(* IEC 61131-3 sources: plc-process-lib/tests/POUs/Suites/FB_AnalogInput_Test, 80 files *)

(* ---- AlarmEventsFailureValueIsRawInput.method.decl.st ---- *)
// Номера и значения событий: udiAlarmIdBase 120 — тревога HH = 120, Failure = 124; значение события HH — rValue_eu
// (95), Failure — сырое rIn (22,5 мА).
METHOD PRIVATE AlarmEventsFailureValueIsRawInput
VAR
    fbTime : FB_FakeTime;         // подменное время
    fbAi   : FB_AnalogInput;      // ФБ под тестом
    stCmd  : ST_AnalogInputCmd;   // команды
    stCfg  : ST_AnalogInputCfg;   // конфигурация
    fbSink : FB_TestSink;         // приёмник событий
    stEv   : ST_AlarmEvent;       // событие
END_VAR

(* ---- At20p5mAIsGood.method.decl.st ---- *)
// Граница 20,5 мА — ещё норма (NE43_MEAS_HIGH_MA: «I > — вне диапазона»): Good, значение 103,125 %.
METHOD PRIVATE At20p5mAIsGood
VAR
    fbTime : FB_FakeTime;         // подменное время
    fbAi   : FB_AnalogInput;      // ФБ под тестом
    stCmd  : ST_AnalogInputCmd;   // команды
    stCfg  : ST_AnalogInputCfg;   // конфигурация
END_VAR

(* ---- At20p7mAIsOutOfSpecification.method.decl.st ---- *)
// 20,7 мА (между 20,5 и 21,0): OverRange, OutOfSpecification, значение — насыщение NE 43 20,5 мА (103,125 %), без
// экстраполяции; выход за диапазон подтверждён — xValid = FALSE (AI-13), бит AI_WRN_OVER_RANGE.
// источник: tools/reference/ai_reference.py, сценарий scale «20,7 мА, шкала 0..100 (насыщение NE 43)».
METHOD PRIVATE At20p7mAIsOutOfSpecification
VAR
    fbTime : FB_FakeTime;         // подменное время
    fbAi   : FB_AnalogInput;      // ФБ под тестом
    stCmd  : ST_AnalogInputCmd;   // команды
    stCfg  : ST_AnalogInputCfg;   // конфигурация
END_VAR

(* ---- At21mAIsFailure.method.decl.st ---- *)
// Граница NE 43 21,0 мА включена в отказ (A-02): FailHigh, Failure, бит AI_FLT_FAIL_HIGH; 20,99 мА — ещё OverRange.
METHOD PRIVATE At21mAIsFailure
VAR
    fbTime : FB_FakeTime;         // подменное время
    fbAi   : FB_AnalogInput;      // ФБ под тестом
    stCmd  : ST_AnalogInputCmd;   // команды
    stCfg  : ST_AnalogInputCfg;   // конфигурация
END_VAR

(* ---- At3p6mAIsFailure.method.decl.st ---- *)
// Граница NE 43 3,6 мА включена в отказ (A-02, сверить с NAMUR NE 43): FailLow, Failure (tFailDelay = 0), бит
// AI_FLT_FAIL_LOW; чуть выше, 3,61 мА — уже UnderRange.
METHOD PRIVATE At3p6mAIsFailure
VAR
    fbTime : FB_FakeTime;         // подменное время
    fbAi   : FB_AnalogInput;      // ФБ под тестом
    stCmd  : ST_AnalogInputCmd;   // команды
    stCfg  : ST_AnalogInputCfg;   // конфигурация
END_VAR

(* ---- At3p7mAIsOutOfSpecification.method.decl.st ---- *)
// 3,7 мА (между 3,6 и 3,8): UnderRange, OutOfSpecification, значение — насыщение NE 43 3,8 мА (-1,25 %), без
// экстраполяции; выход за диапазон подтверждён (tFailDelay = 0) — xValid = FALSE (AI-13), бит AI_WRN_UNDER_RANGE,
// тревога OutOfRange. источник: tools/reference/ai_reference.py, сценарий scale «3,7 мА, шкала 0..100 (насыщение
// NE 43)».
METHOD PRIVATE At3p7mAIsOutOfSpecification
VAR
    fbTime : FB_FakeTime;         // подменное время
    fbAi   : FB_AnalogInput;      // ФБ под тестом
    stCmd  : ST_AnalogInputCmd;   // команды
    stCfg  : ST_AnalogInputCfg;   // конфигурация
    itfAlm : I_Alarm;             // слот тревоги через интерфейс
END_VAR

(* ---- At3p8mAIsGood.method.decl.st ---- *)
// Граница 3,8 мА — уже норма (NE43_MEAS_LOW_MA: «I < — вне диапазона»): Good, значение -1,25 %.
METHOD PRIVATE At3p8mAIsGood
VAR
    fbTime : FB_FakeTime;         // подменное время
    fbAi   : FB_AnalogInput;      // ФБ под тестом
    stCmd  : ST_AnalogInputCmd;   // команды
    stCfg  : ST_AnalogInputCfg;   // конфигурация
END_VAR

(* ---- CfgErrBitsMatchContractMap.method.decl.st ---- *)
// Каждая проверка CheckConfig ставит свой бит wCfgErr (карта 11.5): тип входа вне перечисления, шкала, порядок уставок,
// уставка вне шкалы, гистерезис (< 0 и >= диапазона), отсечка (вне 0…20 %), значение отказа (вне перечисления и NaN),
// приоритет тревоги вне перечисления, шкала отсчётов Raw. Один экземпляр: wCfgErr — результат проверки этого вызова.
METHOD PRIVATE CfgErrBitsMatchContractMap
VAR
    fbTime : FB_FakeTime;         // подменное время
    fbAi   : FB_AnalogInput;      // ФБ под тестом
    stCmd  : ST_AnalogInputCmd;   // команды
    stCfg  : ST_AnalogInputCfg;   // конфигурация
    stBad  : ST_AnalogInputCfg;   // испорченная копия
    uEnum  : U_AiDiTestEnum;      // значение вне строгого перечисления
    uPrio  : U_TestEnumInt;       // приоритет вне перечисления
    uBits  : U_RealBits;          // NaN по битам
END_VAR

(* ---- ChannelFaultSetsFailure.method.decl.st ---- *)
// xChannelFault (диагностика модуля, ошибка обмена) при нормальном токе: ChannelFault, значение удерживается, через
// tFailDelay 2 с — Failure и бит AI_FLT_CHANNEL; после снятия — возврат через те же 2 с.
METHOD PRIVATE ChannelFaultSetsFailure
VAR
    fbTime : FB_FakeTime;         // подменное время
    fbAi   : FB_AnalogInput;      // ФБ под тестом
    stCmd  : ST_AnalogInputCmd;   // команды
    stCfg  : ST_AnalogInputCfg;   // конфигурация
    iStep  : INT;                 // шаг цикла
END_VAR

(* ---- ChannelFaultSetsFailure.method.impl.st ---- *)
coUnit.TEST('AnalogInput_ChannelFault_SetsFailure');

fbAi(itfTime := fbTime, rIn := 12.0, stCmd := stCmd, stCfg := stCfg);   // t0: 50
fbTime.Advance(tStep := T#100MS);
// t1 = t0 + 0,1 с: отказ канала
fbAi(itfTime := fbTime, rIn := 12.0, xChannelFault := TRUE, stCmd := stCmd, stCfg := stCfg);
FOR iStep := 1 TO 19 DO   // t1 + 1,9 с
    fbTime.Advance(tStep := T#100MS);
    fbAi(itfTime := fbTime, rIn := 12.0, xChannelFault := TRUE, stCmd := stCmd, stCfg := stCfg);
END_FOR
AssertTrue(Condition := fbAi.stSts.eSignal = E_AiSignalState.ChannelFault, Message := 'ChannelFault');
AssertFalse(Condition := fbAi.Fault, Message := 'no failure before tFailDelay');
fbTime.Advance(tStep := T#100MS);
fbAi(itfTime := fbTime, rIn := 12.0, xChannelFault := TRUE, stCmd := stCmd, stCfg := stCfg);   // t1 + 2,0 с
AssertTrue(Condition := fbAi.Fault, Message := 'failure after tFailDelay');
AssertEquals_WORD(Expected := GVL_Const.AI_FLT_CHANNEL, Actual := fbAi.stSts.stCommon.wFault, Message := 'CHANNEL bit');
AssertEquals_REAL(Expected := 50.0, Actual := fbAi.rValue_eu, Delta := 1.0E-4, Message := 'value held');
fbTime.Advance(tStep := T#100MS);
fbAi(itfTime := fbTime, rIn := 12.0, xChannelFault := FALSE, stCmd := stCmd, stCfg := stCfg);   // tc: отказ канала снят
FOR iStep := 1 TO 19 DO   // tc + 1,9 с
    fbTime.Advance(tStep := T#100MS);
    fbAi(itfTime := fbTime, rIn := 12.0, xChannelFault := FALSE, stCmd := stCmd, stCfg := stCfg);
END_FOR
AssertTrue(Condition := fbAi.Fault, Message := 'failure kept during return confirmation');
AssertEquals_WORD(Expected := 0, Actual := fbAi.stSts.stCommon.wFault,
                  Message := 'fault bit by current classification');
FOR iStep := 1 TO 1 DO   // tc + 2,0 с
    fbTime.Advance(tStep := T#100MS);
    fbAi(itfTime := fbTime, rIn := 12.0, xChannelFault := FALSE, stCmd := stCmd, stCfg := stCfg);
END_FOR
AssertFalse(Condition := fbAi.Fault, Message := 'failure cleared');

coUnit.TEST_FINISHED();

(* ---- ClampLimitsToRange.method.decl.st ---- *)
// По умолчанию значение экстраполируется (20,4 мА — 102,5 %); с xClamp — ограничено шкалой (100 и 0) с предупреждением
// AI_WRN_CLAMPED. источник: tools/reference/ai_reference.py, сценарии scale «20,4 мА без ограничения», «… с
// ограничением», «3,9 мА с ограничением».
METHOD PRIVATE ClampLimitsToRange
VAR
    fbTime : FB_FakeTime;         // подменное время
    fbAi   : FB_AnalogInput;      // ФБ под тестом
    stCmd  : ST_AnalogInputCmd;   // команды
    stCfg  : ST_AnalogInputCfg;   // конфигурация
END_VAR

(* ---- DefaultCfgFirstCallAutoTypeAndSlots.method.decl.st ---- *)
// Cfg по умолчанию проходит CheckConfig (wCfgErr = 0); после первого вызова — Auto («Измерение»), тип AnalogInput, 6
// слотов тревог, Good, бит DEV_STS_MODE_AUTO; седьмого слота нет; Local не запрашивается.
METHOD PRIVATE DefaultCfgFirstCallAutoTypeAndSlots
VAR
    fbTime : FB_FakeTime;         // подменное время
    fbAi   : FB_AnalogInput;      // ФБ под тестом
    stCmd  : ST_AnalogInputCmd;   // команды
    stCfg  : ST_AnalogInputCfg;   // конфигурация
    itfAlm : I_Alarm;             // слот тревоги через интерфейс
END_VAR

(* ---- EngInputPassesThrough.method.decl.st ---- *)
// Eng (значение уже в инж. ед., Modbus REAL): шкала -50..150, 123,4 — 123,4 (86,7 %); NE 43 не применяется (0 — норма).
// источник: tools/reference/ai_reference.py, сценарий scale «Eng 123,4, шкала -50..150».
METHOD PRIVATE EngInputPassesThrough
VAR
    fbTime : FB_FakeTime;         // подменное время
    fbAi   : FB_AnalogInput;      // ФБ под тестом
    stCmd  : ST_AnalogInputCmd;   // команды
    stCfg  : ST_AnalogInputCfg;   // конфигурация
END_VAR

(* ---- FailureForcesLimitsFalseAndSuppressesLimitAlarms.method.decl.st ---- *)
// H 4,0 активна (4,25 м); обрыв: пока отказ не подтверждён, H держится по удержанному значению, ложного LL (0,5) нет;
// после подтверждения флаги сняты, тревога H — SuppressedByDesign, тревога Failure — ActiveUnack.
METHOD PRIVATE FailureForcesLimitsFalseAndSuppressesLimitAlarms
VAR
    fbTime : FB_FakeTime;         // подменное время
    fbAi   : FB_AnalogInput;      // ФБ под тестом
    stCmd  : ST_AnalogInputCmd;   // команды
    stCfg  : ST_AnalogInputCfg;   // конфигурация
    itfAlm : I_Alarm;             // слот тревоги через интерфейс
    iStep  : INT;                 // шаг цикла
END_VAR

(* ---- FailureForcesLimitsFalseAndSuppressesLimitAlarms.method.impl.st ---- *)
coUnit.TEST('AnalogInput_Failure_ForcesLimitsFalseAndSuppressesLimitAlarms');

stCfg.rRangeHi_eu := 5.0;
SetLimit(stCfgAi := stCfg, uiIdx := E_AiAlarm.H, xEnable := TRUE, rSp_eu := 4.0, rHyst_eu := 0.1, tOnDly := T#0S,
         tOffDly := T#0S);
SetLimit(stCfgAi := stCfg, uiIdx := E_AiAlarm.LL, xEnable := TRUE, rSp_eu := 0.5, rHyst_eu := 0.1, tOnDly := T#0S,
         tOffDly := T#0S);
fbAi(itfTime := fbTime, rIn := 17.6, stCmd := stCmd, stCfg := stCfg);   // t0: 4,25 м
AssertTrue(Condition := fbAi.xH, Message := 'H active before break');
itfAlm := fbAi.GetAlarm(uiIndex := E_AiAlarm.H);
AssertTrue(Condition := itfAlm.State = E_AlarmState.ActiveUnack, Message := 'H alarm active');
fbTime.Advance(tStep := T#100MS);
fbAi(itfTime := fbTime, rIn := 0.0, stCmd := stCmd, stCfg := stCfg);   // t1 = t0 + 0,1 с: обрыв
FOR iStep := 1 TO 19 DO   // t1 + 1,9 с
    fbTime.Advance(tStep := T#100MS);
    fbAi(itfTime := fbTime, rIn := 0.0, stCmd := stCmd, stCfg := stCfg);
END_FOR
AssertTrue(Condition := fbAi.xH, Message := 'H kept on held value while pending');
AssertFalse(Condition := fbAi.xLL, Message := 'no false LL while pending');
fbTime.Advance(tStep := T#100MS);
fbAi(itfTime := fbTime, rIn := 0.0, stCmd := stCmd, stCfg := stCfg);   // t1 + 2,0 с
AssertTrue(Condition := fbAi.Fault, Message := 'failure confirmed');
AssertFalse(Condition := fbAi.xH, Message := 'H forced off');
AssertFalse(Condition := fbAi.xLL, Message := 'LL forced off');
AssertTrue(Condition := itfAlm.State = E_AlarmState.SuppressedByDesign, Message := 'H alarm suppressed');
itfAlm := fbAi.GetAlarm(uiIndex := E_AiAlarm.Failure);
AssertTrue(Condition := itfAlm.State = E_AlarmState.ActiveUnack, Message := 'failure alarm');

coUnit.TEST_FINISHED();

(* ---- FailValueSubstituteUsesCfgValue.method.decl.st ---- *)
// eFailValue = Substitute: до подтверждения отказа держится последнее хорошее значение (25), после — rFailValue_eu =
// 99, xValid = FALSE.
METHOD PRIVATE FailValueSubstituteUsesCfgValue
VAR
    fbTime : FB_FakeTime;         // подменное время
    fbAi   : FB_AnalogInput;      // ФБ под тестом
    stCmd  : ST_AnalogInputCmd;   // команды
    stCfg  : ST_AnalogInputCfg;   // конфигурация
    iStep  : INT;                 // шаг цикла
END_VAR

(* ---- FailValueSubstituteUsesCfgValue.method.impl.st ---- *)
coUnit.TEST('AnalogInput_FailValueSubstitute_UsesCfgValue');

stCfg.eFailValue := E_AiFailValue.Substitute;
stCfg.rFailValue_eu := 99.0;
stCfg.tFailDelay := T#1S;
fbAi(itfTime := fbTime, rIn := 8.0, stCmd := stCmd, stCfg := stCfg);   // t0: 25
fbTime.Advance(tStep := T#100MS);
fbAi(itfTime := fbTime, rIn := 0.0, stCmd := stCmd, stCfg := stCfg);   // t1 = t0 + 0,1 с: обрыв
FOR iStep := 1 TO 9 DO   // t1 + 0,9 с
    fbTime.Advance(tStep := T#100MS);
    fbAi(itfTime := fbTime, rIn := 0.0, stCmd := stCmd, stCfg := stCfg);
END_FOR
AssertEquals_REAL(Expected := 25.0, Actual := fbAi.rValue_eu, Delta := 1.0E-4, Message := 'last good while pending');
AssertTrue(Condition := fbAi.xValid, Message := 'valid while pending');
FOR iStep := 1 TO 1 DO   // t1 + 1,0 с
    fbTime.Advance(tStep := T#100MS);
    fbAi(itfTime := fbTime, rIn := 0.0, stCmd := stCmd, stCfg := stCfg);
END_FOR
AssertTrue(Condition := fbAi.Fault, Message := 'failure confirmed');
AssertEquals_REAL(Expected := 99.0, Actual := fbAi.rValue_eu, Delta := 0.0, Message := 'substitute value from Cfg');
AssertFalse(Condition := fbAi.xValid, Message := 'substitute value is not valid');

coUnit.TEST_FINISHED();

(* ---- FilterIndependentOfCycleTime.method.decl.st ---- *)
// Один и тот же интервал 5 с при T = 10 с: шаг 10 мс (500 вызовов), 250 мс (20 вызовов) и неравномерный 50/150/300 мс
// дают одно значение 39,347 (1 - e^-0,5): фильтр считает по реальному шагу времени. Неявный Эйлер dt/(T + dt) при 250
// мс дал бы 38,97. источник: tools/reference/ai_reference.py, сценарии filter «5 с шагом 10 мс», «… 250 мс», «…
// неравномерно».
METHOD PRIVATE FilterIndependentOfCycleTime
VAR
    fbTimeA : FB_FakeTime;         // время экземпляра A
    fbTimeB : FB_FakeTime;         // время экземпляра B
    fbTimeC : FB_FakeTime;         // время экземпляра C
    fbAiA   : FB_AnalogInput;      // шаг 10 мс
    fbAiB   : FB_AnalogInput;      // шаг 250 мс
    fbAiC   : FB_AnalogInput;      // неравномерный шаг
    stCmdA  : ST_AnalogInputCmd;   // команды A
    stCmdB  : ST_AnalogInputCmd;   // команды B
    stCmdC  : ST_AnalogInputCmd;   // команды C
    stCfg   : ST_AnalogInputCfg;   // конфигурация
    iStep   : INT;                 // шаг цикла
END_VAR

(* ---- FilterIndependentOfCycleTime.method.impl.st ---- *)
coUnit.TEST('AnalogInput_Filter_IndependentOfCycleTime');

stCfg.tFilter := T#10S;
fbAiA(itfTime := fbTimeA, rIn := 4.0, stCmd := stCmdA, stCfg := stCfg);
fbAiB(itfTime := fbTimeB, rIn := 4.0, stCmd := stCmdB, stCfg := stCfg);
fbAiC(itfTime := fbTimeC, rIn := 4.0, stCmd := stCmdC, stCfg := stCfg);
FOR iStep := 1 TO 500 DO
    fbTimeA.Advance(tStep := T#10MS);
    fbAiA(itfTime := fbTimeA, rIn := 20.0, stCmd := stCmdA, stCfg := stCfg);
END_FOR
FOR iStep := 1 TO 20 DO
    fbTimeB.Advance(tStep := T#250MS);
    fbAiB(itfTime := fbTimeB, rIn := 20.0, stCmd := stCmdB, stCfg := stCfg);
END_FOR
FOR iStep := 1 TO 10 DO
    fbTimeC.Advance(tStep := T#50MS);
    fbAiC(itfTime := fbTimeC, rIn := 20.0, stCmd := stCmdC, stCfg := stCfg);
    fbTimeC.Advance(tStep := T#150MS);
    fbAiC(itfTime := fbTimeC, rIn := 20.0, stCmd := stCmdC, stCfg := stCfg);
    fbTimeC.Advance(tStep := T#300MS);
    fbAiC(itfTime := fbTimeC, rIn := 20.0, stCmd := stCmdC, stCfg := stCfg);
END_FOR
AssertEquals_REAL(Expected := 39.34694, Actual := fbAiA.rValue_eu, Delta := 1.0E-3, Message := '10 ms steps');
AssertEquals_REAL(Expected := 39.34694, Actual := fbAiB.rValue_eu, Delta := 1.0E-3, Message := '250 ms steps');
AssertEquals_REAL(Expected := 39.34694, Actual := fbAiC.rValue_eu, Delta := 1.0E-3, Message := 'irregular steps');
AssertEquals_REAL(Expected := fbAiA.rValue_eu, Actual := fbAiB.rValue_eu, Delta := 1.0E-4,
                  Message := 'same result for 10 ms and 250 ms');

coUnit.TEST_FINISHED();

(* ---- FilterOneTimeConstantReaches63Pct.method.decl.st ---- *)
// Фильтр T = 10 с, ступень 0 -> 100 % с шагом 100 мс: в 9,9 с — 62,842, ровно через T — 63,212 (1 - e^-1). источник:
// tools/reference/ai_reference.py, сценарии filter «… 99 шагов по 0,1 с» и «… 100 шагов по 0,1 с».
METHOD PRIVATE FilterOneTimeConstantReaches63Pct
VAR
    fbTime : FB_FakeTime;         // подменное время
    fbAi   : FB_AnalogInput;      // ФБ под тестом
    stCmd  : ST_AnalogInputCmd;   // команды
    stCfg  : ST_AnalogInputCfg;   // конфигурация
    iStep  : INT;                 // шаг цикла
END_VAR

(* ---- FilterOneTimeConstantReaches63Pct.method.impl.st ---- *)
coUnit.TEST('AnalogInput_Filter_OneTimeConstant_Reaches63Pct');

stCfg.tFilter := T#10S;
fbAi(itfTime := fbTime, rIn := 4.0, stCmd := stCmd, stCfg := stCfg);   // t0: фильтр начат с 0
FOR iStep := 1 TO 99 DO   // ступень 100 %, t0 + 9,9 с
    fbTime.Advance(tStep := T#100MS);
    fbAi(itfTime := fbTime, rIn := 20.0, stCmd := stCmd, stCfg := stCfg);
END_FOR
AssertEquals_REAL(Expected := 62.84233, Actual := fbAi.rValue_eu, Delta := 1.0E-3, Message := '62.84 at 9.9 s');
fbTime.Advance(tStep := T#100MS);
fbAi(itfTime := fbTime, rIn := 20.0, stCmd := stCmd, stCfg := stCfg);   // t0 + 10,0 с
AssertEquals_REAL(Expected := 63.21206, Actual := fbAi.rValue_eu, Delta := 1.0E-3, Message := '63.2 % after one T');

coUnit.TEST_FINISHED();

(* ---- GuardBandHighInvalidLimitsKept.method.decl.st ---- *)
// 20,9 мА — верхняя защитная полоса NE 43 (между 20,5 и 21 мА, AI-13): значение — насыщение 20,5 мА, 10,3125 м на
// шкале 0..10 м (1,03125 · 10), без экстраполяции; через tFailDelay — xValid = FALSE, OVER_RANGE, уставка HH (9,5 м)
// остаётся: процесс выше верхнего предела измерения. источник: tools/reference/ai_reference.py, сценарий scale
// «20,9 мА, шкала 0..10 (насыщение NE 43)».
METHOD PRIVATE GuardBandHighInvalidLimitsKept
VAR
    fbTime : FB_FakeTime;         // подменное время
    fbAi   : FB_AnalogInput;      // ФБ под тестом
    stCmd  : ST_AnalogInputCmd;   // команды
    stCfg  : ST_AnalogInputCfg;   // конфигурация
    iStep  : INT;                 // шаг цикла
END_VAR

(* ---- GuardBandHighInvalidLimitsKept.method.impl.st ---- *)
coUnit.TEST('AnalogInput_GuardBandHigh_InvalidLimitsKept');

stCfg.rRangeHi_eu := 10.0;
stCfg.astLimit[E_AiAlarm.HH].xEnable := TRUE;
stCfg.astLimit[E_AiAlarm.HH].rSetpoint_eu := 9.5;
fbAi(itfTime := fbTime, rIn := 12.0, stCmd := stCmd, stCfg := stCfg);                 // t0: 5 м
FOR iStep := 1 TO 21 DO                                                              // t1 + 2,0 с
    fbTime.Advance(tStep := T#100MS);
    fbAi(itfTime := fbTime, rIn := 20.9, stCmd := stCmd, stCfg := stCfg);
END_FOR
AssertEquals_REAL(Expected := 10.3125, Actual := fbAi.rValue_eu, Delta := 1.0E-4,
                  Message := 'no extrapolation above the 20.5 mA saturation');
AssertFalse(Condition := fbAi.xValid, Message := 'confirmed guard band: invalid for control');
AssertEquals_WORD(Expected := GVL_Const.AI_WRN_OVER_RANGE, Actual := fbAi.stSts.stCommon.wWarning,
                  Message := 'over range warning');
AssertEquals_WORD(Expected := 0, Actual := fbAi.stSts.stCommon.wFault, Message := 'no fault bits');
AssertTrue(Condition := fbAi.xHH, Message := 'HH kept');

coUnit.TEST_FINISHED();

(* ---- GuardBandLowInvalidAfterDelay.method.decl.st ---- *)
// 3,61 мА — защитная полоса NE 43 между отказом (<= 3,6) и измерением (>= 3,8 мА): исправный датчик NE 43 так не
// выдаёт, это ток отказа с погрешностью канала или насыщение (AI-13). Значение не экстраполируется ниже насыщения
// 3,8 мА: -0,125 м на шкале 0..10 м (-0,0125 · 10). Пока выход за диапазон не подтверждён (1,9 с) — xValid; через
// tFailDelay = 2 с — xValid = FALSE (ПИД и автоматика по неопределённому значению не управляют), NE 107
// OutOfSpecification, wFault = 0, UNDER_RANGE; уставка LL остаётся (значение не выше насыщения). Норма 12 мА —
// xValid снова через tFailDelay. источник: tools/reference/ai_reference.py, сценарий scale «3,61 мА, шкала 0..10
// (насыщение NE 43)».
METHOD PRIVATE GuardBandLowInvalidAfterDelay
VAR
    fbTime : FB_FakeTime;         // подменное время
    fbAi   : FB_AnalogInput;      // ФБ под тестом
    stCmd  : ST_AnalogInputCmd;   // команды
    stCfg  : ST_AnalogInputCfg;   // конфигурация
    iStep  : INT;                 // шаг цикла
END_VAR

(* ---- GuardBandLowInvalidAfterDelay.method.impl.st ---- *)
coUnit.TEST('AnalogInput_GuardBandLow_InvalidAfterDelay');

stCfg.rRangeHi_eu := 10.0;
stCfg.astLimit[E_AiAlarm.LL].xEnable := TRUE;
stCfg.astLimit[E_AiAlarm.LL].rSetpoint_eu := 0.5;
fbAi(itfTime := fbTime, rIn := 12.0, stCmd := stCmd, stCfg := stCfg);                 // t0: 5 м
FOR iStep := 1 TO 20 DO                                                              // t1 = t0 + 0,1 с … t1 + 1,9 с
    fbTime.Advance(tStep := T#100MS);
    fbAi(itfTime := fbTime, rIn := 3.61, stCmd := stCmd, stCfg := stCfg);
END_FOR
AssertTrue(Condition := fbAi.xValid, Message := 'valid while out of range is unconfirmed (1.9 s)');
AssertEquals_REAL(Expected := -0.125, Actual := fbAi.rValue_eu, Delta := 1.0E-5,
                  Message := 'no extrapolation below the 3.8 mA saturation');
fbTime.Advance(tStep := T#100MS);
fbAi(itfTime := fbTime, rIn := 3.61, stCmd := stCmd, stCfg := stCfg);                  // t1 + 2,0 с
AssertFalse(Condition := fbAi.xValid, Message := 'confirmed guard band: invalid for control');
AssertEquals_REAL(Expected := -0.125, Actual := fbAi.rValue_eu, Delta := 1.0E-5, Message := 'value at saturation');
AssertTrue(Condition := fbAi.Status = E_Ne107Status.OutOfSpecification, Message := 'out of specification, not failure');
AssertEquals_WORD(Expected := 0, Actual := fbAi.stSts.stCommon.wFault, Message := 'no fault bits');
AssertEquals_WORD(Expected := GVL_Const.AI_WRN_UNDER_RANGE, Actual := fbAi.stSts.stCommon.wWarning,
                  Message := 'under range warning');
AssertTrue(Condition := fbAi.xLL, Message := 'LL kept');
FOR iStep := 1 TO 21 DO                                                              // возврат + 2,0 с
    fbTime.Advance(tStep := T#100MS);
    fbAi(itfTime := fbTime, rIn := 12.0, stCmd := stCmd, stCfg := stCfg);
END_FOR
AssertTrue(Condition := fbAi.xValid, Message := 'valid again after tFailDelay in range');
AssertEquals_REAL(Expected := 5.0, Actual := fbAi.rValue_eu, Delta := 1.0E-4, Message := 'measured value');

coUnit.TEST_FINISHED();

(* ---- InvalidRangeAtStartupCheckFunctionSafeValue.method.decl.st ---- *)
// Шкала 10..10 с первого вызова: бит AI_CFG_RANGE, CheckFunction, безопасное значение 0.0, xValid = FALSE, флаги
// уставок FALSE, Available = FALSE; режим — Auto, тип — AnalogInput.
METHOD PRIVATE InvalidRangeAtStartupCheckFunctionSafeValue
VAR
    fbTime : FB_FakeTime;         // подменное время
    fbAi   : FB_AnalogInput;      // ФБ под тестом
    stCmd  : ST_AnalogInputCmd;   // команды
    stCfg  : ST_AnalogInputCfg;   // конфигурация
END_VAR

(* ---- LimitDisabledNeverSets.method.decl.st ---- *)
// Выключенные уставки (HH 10 и LL 90 при значении 50) флаги не взводят ни в одном вызове и не проверяются CheckConfig
// (порядок и шкала — только у включённых).
METHOD PRIVATE LimitDisabledNeverSets
VAR
    fbTime   : FB_FakeTime;         // подменное время
    fbAi     : FB_AnalogInput;      // ФБ под тестом
    stCmd    : ST_AnalogInputCmd;   // команды
    stCfg    : ST_AnalogInputCfg;   // конфигурация
    itfAlm   : I_Alarm;             // слот тревоги через интерфейс
    iStep    : INT;                 // шаг цикла
    xEverSet : BOOL;                // флаг взводился хотя бы раз
END_VAR

(* ---- LimitDisabledNeverSets.method.impl.st ---- *)
coUnit.TEST('AnalogInput_LimitDisabled_NeverSets');

stCfg.eInput := E_AiInputType.Eng;
stCfg.tFailDelay := T#0S;
SetLimit(stCfgAi := stCfg, uiIdx := E_AiAlarm.HH, xEnable := FALSE, rSp_eu := 10.0, rHyst_eu := 0.0, tOnDly := T#0S,
         tOffDly := T#0S);
SetLimit(stCfgAi := stCfg, uiIdx := E_AiAlarm.LL, xEnable := FALSE, rSp_eu := 90.0, rHyst_eu := 0.0, tOnDly := T#0S,
         tOffDly := T#0S);
fbAi(itfTime := fbTime, rIn := 50.0, stCmd := stCmd, stCfg := stCfg);
FOR iStep := 1 TO 10 DO
    fbTime.Advance(tStep := T#100MS);
    fbAi(itfTime := fbTime, rIn := 50.0, stCmd := stCmd, stCfg := stCfg);
    xEverSet := xEverSet OR fbAi.xHH OR fbAi.xLL;
END_FOR
AssertFalse(Condition := xEverSet, Message := 'disabled limits never set');
AssertEquals_WORD(Expected := 0, Actual := fbAi.stSts.stCommon.wCfgErr, Message := 'disabled limits are not checked');
itfAlm := fbAi.GetAlarm(uiIndex := E_AiAlarm.HH);
AssertTrue(Condition := itfAlm.State = E_AlarmState.Normal, Message := 'HH alarm normal');

coUnit.TEST_FINISHED();

(* ---- LimitHHOnDelayShortExcursionIgnored.method.decl.st ---- *)
// HH 90 с задержкой срабатывания 3 с: выброс 2,9 с флаг не взводит; устойчивое превышение — флаг ровно через 3,0 с.
METHOD PRIVATE LimitHHOnDelayShortExcursionIgnored
VAR
    fbTime  : FB_FakeTime;         // подменное время
    fbAi    : FB_AnalogInput;      // ФБ под тестом
    stCmd   : ST_AnalogInputCmd;   // команды
    stCfg   : ST_AnalogInputCfg;   // конфигурация
    iStep   : INT;                 // шаг цикла
    xEverHH : BOOL;                // HH взводился хотя бы раз
END_VAR

(* ---- LimitHHOnDelayShortExcursionIgnored.method.impl.st ---- *)
coUnit.TEST('AnalogInput_LimitHH_OnDelay_ShortExcursionIgnored');

stCfg.eInput := E_AiInputType.Eng;
stCfg.tFailDelay := T#0S;
SetLimit(stCfgAi := stCfg, uiIdx := E_AiAlarm.HH, xEnable := TRUE, rSp_eu := 90.0, rHyst_eu := 1.0, tOnDly := T#3S,
         tOffDly := T#0S);
fbAi(itfTime := fbTime, rIn := 95.0, stCmd := stCmd, stCfg := stCfg);   // t0: выброс
FOR iStep := 1 TO 29 DO                                           // t0 + 2,9 с
    fbTime.Advance(tStep := T#100MS);
    fbAi(itfTime := fbTime, rIn := 95.0, stCmd := stCmd, stCfg := stCfg);
    xEverHH := xEverHH OR fbAi.xHH;
END_FOR
fbTime.Advance(tStep := T#100MS);
fbAi(itfTime := fbTime, rIn := 85.0, stCmd := stCmd, stCfg := stCfg);   // t0 + 3,0 с: выброс кончился
xEverHH := xEverHH OR fbAi.xHH;
AssertFalse(Condition := xEverHH, Message := 'excursion shorter than on-delay ignored');
fbTime.Advance(tStep := T#100MS);
fbAi(itfTime := fbTime, rIn := 95.0, stCmd := stCmd, stCfg := stCfg);   // t1
FOR iStep := 1 TO 29 DO   // t1 + 2,9 с
    fbTime.Advance(tStep := T#100MS);
    fbAi(itfTime := fbTime, rIn := 95.0, stCmd := stCmd, stCfg := stCfg);
END_FOR
AssertFalse(Condition := fbAi.xHH, Message := 'no HH at t1 + 2.9 s');
fbTime.Advance(tStep := T#100MS);
fbAi(itfTime := fbTime, rIn := 95.0, stCmd := stCmd, stCfg := stCfg);   // t1 + 3,0 с
AssertTrue(Condition := fbAi.xHH, Message := 'HH exactly at t1 + 3.0 s');

coUnit.TEST_FINISHED();

(* ---- LimitHHysteresisClearsBelowSpMinusHyst.method.decl.st ---- *)
// Уставка H 80, гистерезис 2 (вход Eng 0..100): 79,9 — нет; 80,0 — да (граница включена); 78,0 — ещё да; 77,9 — снят.
// Тревога H — ActiveUnack, бит AI_STS_H.
METHOD PRIVATE LimitHHysteresisClearsBelowSpMinusHyst
VAR
    fbTime : FB_FakeTime;         // подменное время
    fbAi   : FB_AnalogInput;      // ФБ под тестом
    stCmd  : ST_AnalogInputCmd;   // команды
    stCfg  : ST_AnalogInputCfg;   // конфигурация
    itfAlm : I_Alarm;             // слот тревоги через интерфейс
END_VAR

(* ---- LimitLHysteresisClearsAboveSpPlusHyst.method.decl.st ---- *)
// Уставка L 20, гистерезис 2: 20,1 — нет; 20,0 — да; 22,0 — ещё да; 22,1 — снят.
METHOD PRIVATE LimitLHysteresisClearsAboveSpPlusHyst
VAR
    fbTime : FB_FakeTime;         // подменное время
    fbAi   : FB_AnalogInput;      // ФБ под тестом
    stCmd  : ST_AnalogInputCmd;   // команды
    stCfg  : ST_AnalogInputCfg;   // конфигурация
END_VAR

(* ---- LimitOffDelayHoldsFlag.method.decl.st ---- *)
// H 80 с задержкой снятия 2 с: значение ушло ниже уставки — флаг держится 1,9 с, снимается в 2,0 с.
METHOD PRIVATE LimitOffDelayHoldsFlag
VAR
    fbTime : FB_FakeTime;         // подменное время
    fbAi   : FB_AnalogInput;      // ФБ под тестом
    stCmd  : ST_AnalogInputCmd;   // команды
    stCfg  : ST_AnalogInputCfg;   // конфигурация
    iStep  : INT;                 // шаг цикла
END_VAR

(* ---- LimitOffDelayHoldsFlag.method.impl.st ---- *)
coUnit.TEST('AnalogInput_LimitOffDelay_HoldsFlag');

stCfg.eInput := E_AiInputType.Eng;
stCfg.tFailDelay := T#0S;
SetLimit(stCfgAi := stCfg, uiIdx := E_AiAlarm.H, xEnable := TRUE, rSp_eu := 80.0, rHyst_eu := 0.0, tOnDly := T#0S,
         tOffDly := T#2S);
fbAi(itfTime := fbTime, rIn := 85.0, stCmd := stCmd, stCfg := stCfg);
AssertTrue(Condition := fbAi.xH, Message := 'H set');
fbTime.Advance(tStep := T#100MS);
fbAi(itfTime := fbTime, rIn := 70.0, stCmd := stCmd, stCfg := stCfg);   // t1: ниже уставки
FOR iStep := 1 TO 19 DO   // t1 + 1,9 с
    fbTime.Advance(tStep := T#100MS);
    fbAi(itfTime := fbTime, rIn := 70.0, stCmd := stCmd, stCfg := stCfg);
END_FOR
AssertTrue(Condition := fbAi.xH, Message := 'H held by off-delay');
fbTime.Advance(tStep := T#100MS);
fbAi(itfTime := fbTime, rIn := 70.0, stCmd := stCmd, stCfg := stCfg);   // t1 + 2,0 с
AssertFalse(Condition := fbAi.xH, Message := 'H cleared after off-delay');

coUnit.TEST_FINISHED();

(* ---- LimitOrderInvalidAtRuntimeKeepsLastValidCfg.method.decl.st ---- *)
// В работе HH испорчена (70 < H 80): бит AI_CFG_LIMIT_ORDER, CheckFunction, но логика работает по последней корректной
// Cfg (HH 90): 85 — только H, 95 — HH; значение пригодно. Исправление Cfg снимает CheckFunction.
METHOD PRIVATE LimitOrderInvalidAtRuntimeKeepsLastValidCfg
VAR
    fbTime : FB_FakeTime;         // подменное время
    fbAi   : FB_AnalogInput;      // ФБ под тестом
    stCmd  : ST_AnalogInputCmd;   // команды
    stCfg  : ST_AnalogInputCfg;   // конфигурация
END_VAR

(* ---- LimitsOnFailEvaluatesFailValue.method.decl.st ---- *)
// xLimitsOnFail = TRUE и Substitute 95: после подтверждения отказа уставки считаются по значению отказа — HH (90)
// взводится, тревога HH не подавлена (ActiveUnack). Так проектировщик задаёт безопасную реакцию на отказ датчика.
METHOD PRIVATE LimitsOnFailEvaluatesFailValue
VAR
    fbTime : FB_FakeTime;         // подменное время
    fbAi   : FB_AnalogInput;      // ФБ под тестом
    stCmd  : ST_AnalogInputCmd;   // команды
    stCfg  : ST_AnalogInputCfg;   // конфигурация
    itfAlm : I_Alarm;             // слот тревоги через интерфейс
    iStep  : INT;                 // шаг цикла
END_VAR

(* ---- LimitsOnFailEvaluatesFailValue.method.impl.st ---- *)
coUnit.TEST('AnalogInput_LimitsOnFail_EvaluatesFailValue');

stCfg.eFailValue := E_AiFailValue.Substitute;
stCfg.rFailValue_eu := 95.0;
stCfg.xLimitsOnFail := TRUE;
stCfg.tFailDelay := T#1S;
SetLimit(stCfgAi := stCfg, uiIdx := E_AiAlarm.HH, xEnable := TRUE, rSp_eu := 90.0, rHyst_eu := 1.0, tOnDly := T#0S,
         tOffDly := T#0S);
fbAi(itfTime := fbTime, rIn := 12.0, stCmd := stCmd, stCfg := stCfg);   // t0: 50
AssertFalse(Condition := fbAi.xHH, Message := 'no HH at 50');
FOR iStep := 1 TO 11 DO   // обрыв с t0 + 0,1 с, t0 + 1,1 с
    fbTime.Advance(tStep := T#100MS);
    fbAi(itfTime := fbTime, rIn := 0.0, stCmd := stCmd, stCfg := stCfg);
END_FOR
AssertTrue(Condition := fbAi.Fault, Message := 'failure confirmed');
AssertEquals_REAL(Expected := 95.0, Actual := fbAi.rValue_eu, Delta := 0.0, Message := 'fail value');
AssertTrue(Condition := fbAi.xHH, Message := 'HH evaluated on fail value');
itfAlm := fbAi.GetAlarm(uiIndex := E_AiAlarm.HH);
AssertTrue(Condition := itfAlm.State = E_AlarmState.ActiveUnack, Message := 'HH alarm not suppressed');

coUnit.TEST_FINISHED();

(* ---- LowCutBelowCutReturnsZero.method.decl.st ---- *)
// Отсечка 5 % после корня: 0,2 % перепада (корень 4,47 %) — 0 и бит AI_STS_LOW_CUT; 1 % перепада (корень 10 %) —
// 9,999995 без бита. Без корня отсечка тоже действует: 2,5 % при отсечке 3 % — 0. Граница: отсечка — при
// x·100 < rLowCut_pct, ровно 12,5 % при отсечке 12,5 % не срезается. источник:
// tools/reference/ai_reference.py, сценарии scale «корень: 4,032 мА», «корень: 4,16 мА», «без корня: 4,4 мА»,
// «без корня: 6 мА (12,5 %), отсечка 12,5 %».
METHOD PRIVATE LowCutBelowCutReturnsZero
VAR
    fbTime : FB_FakeTime;         // подменное время
    fbAi   : FB_AnalogInput;      // ФБ под тестом
    stCmd  : ST_AnalogInputCmd;   // команды
    stCfg  : ST_AnalogInputCfg;   // конфигурация
END_VAR

(* ---- NaNInputTreatedAsFailure.method.decl.st ---- *)
// NaN на входе (например, ошибка обмена REAL): NotFinite, значение удерживается до подтверждения (tFailDelay 1 с),
// затем Failure и бит AI_FLT_NOT_FINITE; +Inf и 1E31 (больше REAL_SANE_MAX) — тоже NotFinite. После возврата значение
// конечно и равно новому: NaN не попал в фильтр.
METHOD PRIVATE NaNInputTreatedAsFailure
VAR
    fbTime : FB_FakeTime;         // подменное время
    fbAi   : FB_AnalogInput;      // ФБ под тестом
    stCmd  : ST_AnalogInputCmd;   // команды
    stCfg  : ST_AnalogInputCfg;   // конфигурация
    iStep  : INT;                 // шаг цикла
    uBits  : U_RealBits;          // NaN и Inf по битам IEEE 754
END_VAR

(* ---- NaNInputTreatedAsFailure.method.impl.st ---- *)
coUnit.TEST('AnalogInput_NaNInput_TreatedAsFailure');

stCfg.tFailDelay := T#1S;
stCfg.tFilter := T#5S;
fbAi(itfTime := fbTime, rIn := 12.0, stCmd := stCmd, stCfg := stCfg);   // t0: 50
uBits.dwValue := 16#7FC00000;                                     // тихий NaN
fbTime.Advance(tStep := T#100MS);
fbAi(itfTime := fbTime, rIn := uBits.rValue, stCmd := stCmd, stCfg := stCfg);   // t1 = t0 + 0,1 с
FOR iStep := 1 TO 9 DO   // t1 + 0,9 с
    fbTime.Advance(tStep := T#100MS);
    fbAi(itfTime := fbTime, rIn := uBits.rValue, stCmd := stCmd, stCfg := stCfg);
END_FOR
AssertTrue(Condition := fbAi.stSts.eSignal = E_AiSignalState.NotFinite, Message := 'NaN is NotFinite');
AssertFalse(Condition := fbAi.Fault, Message := 'no failure before tFailDelay');
// AssertEquals_REAL пропускает NaN (ABS(NaN) > Delta = FALSE): конечность проверяется отдельно
AssertTrue(Condition := F_IsFinite(rIn := fbAi.rValue_eu) AND F_IsFinite(rIn := fbAi.rValue_pct),
           Message := 'NaN input: value finite');
AssertTrue(Condition := F_IsFinite(rIn := stCmd.rSubstValue_eu), Message := 'NaN input: substitution tracking finite');
AssertEquals_REAL(Expected := 50.0, Actual := fbAi.rValue_eu, Delta := 1.0E-4, Message := 'value held, not NaN');
fbTime.Advance(tStep := T#100MS);
fbAi(itfTime := fbTime, rIn := uBits.rValue, stCmd := stCmd, stCfg := stCfg);   // t1 + 1,0 с
AssertTrue(Condition := fbAi.Status = E_Ne107Status.Failure, Message := 'failure after tFailDelay');
AssertEquals_WORD(Expected := GVL_Const.AI_FLT_NOT_FINITE, Actual := fbAi.stSts.stCommon.wFault,
                  Message := 'NOT_FINITE fault bit');
uBits.dwValue := 16#7F800000;                                     // +Inf
fbTime.Advance(tStep := T#100MS);
fbAi(itfTime := fbTime, rIn := uBits.rValue, stCmd := stCmd, stCfg := stCfg);
AssertTrue(Condition := fbAi.stSts.eSignal = E_AiSignalState.NotFinite, Message := '+Inf is NotFinite');
AssertTrue(Condition := F_IsFinite(rIn := fbAi.rValue_eu) AND F_IsFinite(rIn := fbAi.rValue_pct),
           Message := '+Inf input: value finite');
fbTime.Advance(tStep := T#100MS);
fbAi(itfTime := fbTime, rIn := 1.0E31, stCmd := stCmd, stCfg := stCfg);
AssertTrue(Condition := fbAi.stSts.eSignal = E_AiSignalState.NotFinite, Message := 'above REAL_SANE_MAX is NotFinite');
fbTime.Advance(tStep := T#100MS);
fbAi(itfTime := fbTime, rIn := 16.0, stCmd := stCmd, stCfg := stCfg);   // tr: сигнал вернулся, 75
FOR iStep := 1 TO 10 DO   // tr + 1,0 с
    fbTime.Advance(tStep := T#100MS);
    fbAi(itfTime := fbTime, rIn := 16.0, stCmd := stCmd, stCfg := stCfg);
END_FOR
AssertFalse(Condition := fbAi.Fault, Message := 'failure cleared');
AssertTrue(Condition := F_IsFinite(rIn := fbAi.rValue_eu), Message := 'value is finite');
AssertEquals_REAL(Expected := 75.0, Actual := fbAi.rValue_eu, Delta := 1.0E-3,
                  Message := 'NaN did not enter the filter');

coUnit.TEST_FINISHED();

(* ---- Norm01NoNe43Check.method.decl.st ---- *)
// Norm01 (0–10 В и т. п.): NE 43 не применяется — rIn = -0,03 даёт экстраполяцию -3 % без отказа и выхода за диапазон
// даже при tFailDelay = 0; 1,5 — 150. источник: tools/reference/ai_reference.py, сценарии scale «Norm01 -0,03» и
// «Norm01 0,7».
METHOD PRIVATE Norm01NoNe43Check
VAR
    fbTime : FB_FakeTime;         // подменное время
    fbAi   : FB_AnalogInput;      // ФБ под тестом
    stCmd  : ST_AnalogInputCmd;   // команды
    stCfg  : ST_AnalogInputCfg;   // конфигурация
END_VAR

(* ---- Norm420ScalesLikeMilliamps.method.decl.st ---- *)
// Norm420: rIn 0..1 = 4..20 мА. 0,5 даёт то же, что 12 мА на соседнем экземпляре (7,0 на шкале 2..12); NE 43 — по
// пересчёту I = 4 + 16·rIn: -0,05 (3,2 мА) — FailLow, 1,0625 (21 мА) — FailHigh. источник:
// tools/reference/ai_reference.py, сценарий scale «Norm420 0,5, шкала 2..12».
METHOD PRIVATE Norm420ScalesLikeMilliamps
VAR
    fbTime  : FB_FakeTime;         // подменное время
    fbAi    : FB_AnalogInput;      // ФБ под тестом
    fbMa    : FB_AnalogInput;      // тот же вход в мА
    stCmd   : ST_AnalogInputCmd;   // команды
    stCmdMa : ST_AnalogInputCmd;   // команды экземпляра в мА
    stCfg   : ST_AnalogInputCfg;   // конфигурация
    stCfgMa : ST_AnalogInputCfg;   // конфигурация экземпляра в мА
END_VAR

(* ---- OosExitWithBrokenSignalInvalidAtOnce.method.decl.st ---- *)
// Выход из OutOfService с уже оборванной линией (датчик меняли «в ремонте», линию ещё не подключили):
// последнее хорошее значение — до вывода из работы, его возраст неизвестен. Удерживать его как годное
// на время подтверждения нельзя: значение сразу негодно, уставки по нему не считаются (как AI-2 при
// старте ПЛК), отказ — через tFailDelay. Шкала 0..5 м: 17,6 мА = 4,25 м (H 4,0), 16 мА = 3,75 м.
METHOD PRIVATE OosExitWithBrokenSignalInvalidAtOnce
VAR
    fbTime : FB_FakeTime;         // подменное время
    fbAi   : FB_AnalogInput;      // ФБ под тестом
    stCmd  : ST_AnalogInputCmd;   // команды
    stCfg  : ST_AnalogInputCfg;   // конфигурация
    iStep  : INT;                 // шаг цикла
END_VAR

(* ---- OosExitWithBrokenSignalInvalidAtOnce.method.impl.st ---- *)
coUnit.TEST('AnalogInput_OosExitWithBrokenSignal_InvalidAtOnce');

stCfg.rRangeHi_eu := 5.0;
SetLimit(stCfgAi := stCfg, uiIdx := E_AiAlarm.H, xEnable := TRUE, rSp_eu := 4.0, rHyst_eu := 0.1, tOnDly := T#0S,
         tOffDly := T#0S);
SetLimit(stCfgAi := stCfg, uiIdx := E_AiAlarm.LL, xEnable := TRUE, rSp_eu := 0.5, rHyst_eu := 0.1, tOnDly := T#0S,
         tOffDly := T#0S);
fbAi(itfTime := fbTime, rIn := 17.6, stCmd := stCmd, stCfg := stCfg);   // t0: 4,25 м, H
AssertTrue(Condition := fbAi.xH, Message := 'H before OOS');
stCmd.stCommon.xSetOos := TRUE;
fbTime.Advance(tStep := T#100MS);
fbAi(itfTime := fbTime, rIn := 17.6, stCmd := stCmd, stCfg := stCfg);   // вывод из работы
FOR iStep := 1 TO 10 DO   // в ремонте: линия оборвана 10 с
    fbTime.Advance(tStep := T#1000MS);
    fbAi(itfTime := fbTime, rIn := 0.0, stCmd := stCmd, stCfg := stCfg);
END_FOR
AssertTrue(Condition := fbAi.Status = E_Ne107Status.CheckFunction, Message := 'no failure in OOS');
stCmd.stCommon.xSetAuto := TRUE;
fbTime.Advance(tStep := T#100MS);
fbAi(itfTime := fbTime, rIn := 0.0, stCmd := stCmd, stCfg := stCfg);    // te: в работу, линия ещё оборвана
AssertTrue(Condition := fbAi.Mode = E_DeviceMode.Auto, Message := 'back in service');
AssertFalse(Condition := fbAi.xValid, Message := 'stale value from before OOS is not valid');
AssertFalse(Condition := fbAi.xH, Message := 'no H from the stale value');
AssertFalse(Condition := fbAi.xLL, Message := 'no false LL');
AssertEquals_REAL(Expected := 4.25, Actual := fbAi.rValue_eu, Delta := 1.0E-5, Message := 'HoldLast keeps held value');
AssertTrue(Condition := (fbAi.stSts.stCommon.wStatus AND GVL_Const.AI_STS_FAIL_PENDING) = 0,
           Message := 'no pending bit: value is not held as valid');
AssertFalse(Condition := fbAi.Fault, Message := 'failure not yet confirmed');
FOR iStep := 1 TO 20 DO   // te + 2,0 с
    fbTime.Advance(tStep := T#100MS);
    fbAi(itfTime := fbTime, rIn := 0.0, stCmd := stCmd, stCfg := stCfg);
END_FOR
AssertTrue(Condition := fbAi.Fault, Message := 'failure after tFailDelay');
FOR iStep := 1 TO 21 DO   // сигнал вернулся, + 2,1 с
    fbTime.Advance(tStep := T#100MS);
    fbAi(itfTime := fbTime, rIn := 16.0, stCmd := stCmd, stCfg := stCfg);
END_FOR
AssertFalse(Condition := fbAi.Fault, Message := 'failure cleared');
AssertTrue(Condition := fbAi.xValid, Message := 'valid with the new measurement');
AssertEquals_REAL(Expected := 3.75, Actual := fbAi.rValue_eu, Delta := 1.0E-5, Message := 'measured value');

coUnit.TEST_FINISHED();

(* ---- OutOfServiceHoldsValueInvalid.method.decl.st ---- *)
// OutOfService: значение удерживается (50 при 16 мА на входе), xValid = FALSE, CheckFunction, флаги уставок сняты, все
// слоты OutOfService; обрыв в OOS не даёт Failure (сигнал не контролируется); слежение пишет удерживаемое значение в
// rSubstValue_eu и в OOS (правило 2.1, AI-10). Выход («Измерение») — измеренное значение 75.
METHOD PRIVATE OutOfServiceHoldsValueInvalid
VAR
    fbTime : FB_FakeTime;         // подменное время
    fbAi   : FB_AnalogInput;      // ФБ под тестом
    stCmd  : ST_AnalogInputCmd;   // команды
    stCfg  : ST_AnalogInputCfg;   // конфигурация
    itfAlm : I_Alarm;             // слот тревоги через интерфейс
    iStep  : INT;                 // шаг цикла
END_VAR

(* ---- OutOfServiceHoldsValueInvalid.method.impl.st ---- *)
coUnit.TEST('AnalogInput_OutOfService_HoldsValueInvalid');

SetLimit(stCfgAi := stCfg, uiIdx := E_AiAlarm.H, xEnable := TRUE, rSp_eu := 40.0, rHyst_eu := 1.0, tOnDly := T#0S,
         tOffDly := T#0S);
fbAi(itfTime := fbTime, rIn := 12.0, stCmd := stCmd, stCfg := stCfg);   // Auto: 50, H
AssertTrue(Condition := fbAi.xH, Message := 'H before OOS');
stCmd.stCommon.xSetOos := TRUE;
fbTime.Advance(tStep := T#100MS);
fbAi(itfTime := fbTime, rIn := 16.0, stCmd := stCmd, stCfg := stCfg);
AssertTrue(Condition := fbAi.Mode = E_DeviceMode.OutOfService, Message := 'out of service');
AssertEquals_REAL(Expected := 50.0, Actual := fbAi.rValue_eu, Delta := 1.0E-4, Message := 'value held');
AssertFalse(Condition := fbAi.xValid, Message := 'invalid in OOS');
AssertTrue(Condition := fbAi.Status = E_Ne107Status.CheckFunction, Message := 'CheckFunction');
AssertFalse(Condition := fbAi.xH, Message := 'limits off in OOS');
itfAlm := fbAi.GetAlarm(uiIndex := E_AiAlarm.H);
AssertTrue(Condition := itfAlm.State = E_AlarmState.OutOfService, Message := 'H slot out of service');
itfAlm := fbAi.GetAlarm(uiIndex := E_AiAlarm.Failure);
AssertTrue(Condition := itfAlm.State = E_AlarmState.OutOfService, Message := 'failure slot out of service');
stCmd.rSubstValue_eu := 7.0;   // оператор пишет поле подмены в OOS
FOR iStep := 1 TO 30 DO   // обрыв в OOS, 3 с
    fbTime.Advance(tStep := T#100MS);
    fbAi(itfTime := fbTime, rIn := 0.0, stCmd := stCmd, stCfg := stCfg);
END_FOR
AssertTrue(Condition := fbAi.Status = E_Ne107Status.CheckFunction, Message := 'no failure in OOS');
AssertEquals_REAL(Expected := 50.0, Actual := stCmd.rSubstValue_eu, Delta := 0.0,
                  Message := 'held value tracked into rSubstValue_eu in OOS');
stCmd.stCommon.xSetAuto := TRUE;
fbTime.Advance(tStep := T#100MS);
fbAi(itfTime := fbTime, rIn := 16.0, stCmd := stCmd, stCfg := stCfg);
AssertTrue(Condition := fbAi.Mode = E_DeviceMode.Auto, Message := 'back in service');
AssertEquals_REAL(Expected := 75.0, Actual := fbAi.rValue_eu, Delta := 1.0E-4, Message := 'measured after OOS');
AssertTrue(Condition := fbAi.xValid, Message := 'valid after OOS');

coUnit.TEST_FINISHED();

(* ---- RawInputScalesCounts.method.decl.st ---- *)
// Raw (целое из Modbus): отсчёты 2000..10000 — шкала 0..16 бар; 6000 — 8,0; 1000 — экстраполяция -2,0; NE 43 не
// применяется, Cfg корректна. источник: tools/reference/ai_reference.py, сценарии scale «Raw 6000» и «Raw 1000».
METHOD PRIVATE RawInputScalesCounts
VAR
    fbTime : FB_FakeTime;         // подменное время
    fbAi   : FB_AnalogInput;      // ФБ под тестом
    stCmd  : ST_AnalogInputCmd;   // команды
    stCfg  : ST_AnalogInputCfg;   // конфигурация
END_VAR

(* ---- RawRangeUnsetCfgErrBit8.method.decl.st ---- *)
// Raw с не заданной шкалой отсчётов (умолчания 0/0): бит 8 wCfgErr (AI_CFG_RAW_RANGE) и только он, CheckFunction,
// безопасное значение 0.0, xValid = FALSE, Available = FALSE. После задания шкалы отсчётов Cfg принимается: 5000 из
// 0..10000 — 50 % шкалы 0..100.
METHOD PRIVATE RawRangeUnsetCfgErrBit8
VAR
    fbTime : FB_FakeTime;         // подменное время
    fbAi   : FB_AnalogInput;      // ФБ под тестом
    stCmd  : ST_AnalogInputCmd;   // команды
    stCfg  : ST_AnalogInputCfg;   // конфигурация
END_VAR

(* ---- ResetCmdAcceptedAndAcksAlarms.method.decl.st ---- *)
// Фиксируемых отказов у AI нет, но xReset — команда: результат Accepted, uiCmdSeq + 1, бит сброшен; неквитированная
// тревога Failure (RtnUnack после возврата сигнала) квитируется — Normal.
METHOD PRIVATE ResetCmdAcceptedAndAcksAlarms
VAR
    fbTime : FB_FakeTime;         // подменное время
    fbAi   : FB_AnalogInput;      // ФБ под тестом
    stCmd  : ST_AnalogInputCmd;   // команды
    stCfg  : ST_AnalogInputCfg;   // конфигурация
    itfAlm : I_Alarm;             // слот тревоги через интерфейс
    uiSeq  : UINT;                // номер команды до сброса
END_VAR

(* ---- Scale12mAReturnsMidRange.method.decl.st ---- *)
// Шкала 2..12: 12 мА — середина шкалы 7,0 (50 %); сырое значение в stSts.rIn. источник:
// tools/reference/ai_reference.py, сценарий scale «12 мА, шкала 2..12».
METHOD PRIVATE Scale12mAReturnsMidRange
VAR
    fbTime : FB_FakeTime;         // подменное время
    fbAi   : FB_AnalogInput;      // ФБ под тестом
    stCmd  : ST_AnalogInputCmd;   // команды
    stCfg  : ST_AnalogInputCfg;   // конфигурация
END_VAR

(* ---- Scale20mAReturnsRangeHi.method.decl.st ---- *)
// Шкала 2..12: 20 мА — конец шкалы 12,0 (100 %). источник: tools/reference/ai_reference.py, сценарий scale «20 мА,
// шкала 2..12».
METHOD PRIVATE Scale20mAReturnsRangeHi
VAR
    fbTime : FB_FakeTime;         // подменное время
    fbAi   : FB_AnalogInput;      // ФБ под тестом
    stCmd  : ST_AnalogInputCmd;   // команды
    stCfg  : ST_AnalogInputCfg;   // конфигурация
END_VAR

(* ---- Scale4mAReturnsRangeLo.method.decl.st ---- *)
// Шкала 2..12: 4 мА — начало шкалы 2,0 (0 %), сигнал в норме, значение пригодно, NE 107 Good. источник:
// tools/reference/ai_reference.py, сценарий scale «4 мА, шкала 2..12».
METHOD PRIVATE Scale4mAReturnsRangeLo
VAR
    fbTime : FB_FakeTime;         // подменное время
    fbAi   : FB_AnalogInput;      // ФБ под тестом
    stCmd  : ST_AnalogInputCmd;   // команды
    stCfg  : ST_AnalogInputCfg;   // конфигурация
END_VAR

(* ---- SetAlarmPriority.method.decl.st ---- *)
// Помощник: приоритет слота тревоги uiSlot в Cfg входа (копия элемента, как SetLimit)
METHOD PRIVATE SetAlarmPriority
VAR_IN_OUT
    stCfgAi : ST_AnalogInputCfg;   // конфигурация входа
END_VAR
VAR_INPUT
    uiSlot    : UINT;              // слот: E_AiAlarm
    ePriority : E_AlarmPriority;   // приоритет
END_VAR
VAR
    stSlot : ST_AlarmCfg;          // копия слота
END_VAR

(* ---- SetLimit.method.decl.st ---- *)
// Помощник: уставка uiIdx (E_AiAlarm.HH, H, L, LL) в Cfg входа (через копию элемента)
METHOD PRIVATE SetLimit
VAR_IN_OUT
    stCfgAi : ST_AnalogInputCfg;   // конфигурация входа
END_VAR
VAR_INPUT
    uiIdx    : UINT;               // уставка: E_AiAlarm.HH, H, L, LL
    xEnable  : BOOL;               // уставка включена
    rSp_eu   : REAL;               // значение уставки, инж. ед.
    rHyst_eu : REAL;               // гистерезис, инж. ед.
    tOnDly   : TIME;               // задержка срабатывания
    tOffDly  : TIME;               // задержка снятия
END_VAR
VAR
    stLim : ST_AiLimitCfg;         // копия уставки
END_VAR

(* ---- ShortGlitchFilterKeptNoFalseLimit.method.decl.st ---- *)
// Короткий провал сигнала (один вызов с отказом канала, ошибка обмена Modbus): отказ не подтверждён, значение
// удерживается, фильтр заморожен и после провала продолжает с прежнего состояния (AI-12). Фильтр 10 с,
// ступень 50 -> 75, HH 70 без задержки: до провала (1 с) 52,379, через вызов после провала 52,604, HH нет.
// Сброс фильтра выдал бы мгновенное 75 и ложный HH. источник: tools/reference/ai_reference.py, сценарии filter
// «ступень 50 -> 75, T = 10 с, 1 с до провала» и «… провал 0,1 с, фильтр заморожен».
METHOD PRIVATE ShortGlitchFilterKeptNoFalseLimit
VAR
    fbTime  : FB_FakeTime;         // подменное время
    fbAi    : FB_AnalogInput;      // ФБ под тестом
    stCmd   : ST_AnalogInputCmd;   // команды
    stCfg   : ST_AnalogInputCfg;   // конфигурация
    iStep   : INT;                 // шаг цикла
    xEverHH : BOOL;                // HH взводился хотя бы раз
END_VAR

(* ---- ShortGlitchFilterKeptNoFalseLimit.method.impl.st ---- *)
coUnit.TEST('AnalogInput_ShortGlitch_FilterKeptNoFalseLimit');

stCfg.tFilter := T#10S;
SetLimit(stCfgAi := stCfg, uiIdx := E_AiAlarm.HH, xEnable := TRUE, rSp_eu := 70.0, rHyst_eu := 1.0, tOnDly := T#0S,
         tOffDly := T#0S);
fbAi(itfTime := fbTime, rIn := 12.0, stCmd := stCmd, stCfg := stCfg);   // t0: фильтр начат с 50
FOR iStep := 1 TO 10 DO   // ступень 75, t0 + 1,0 с
    fbTime.Advance(tStep := T#100MS);
    fbAi(itfTime := fbTime, rIn := 16.0, stCmd := stCmd, stCfg := stCfg);
END_FOR
AssertEquals_REAL(Expected := 52.37906, Actual := fbAi.rValue_eu, Delta := 1.0E-3, Message := 'filtered before glitch');
fbTime.Advance(tStep := T#100MS);
fbAi(itfTime := fbTime, rIn := 16.0, xChannelFault := TRUE, stCmd := stCmd, stCfg := stCfg);   // провал
AssertEquals_REAL(Expected := 52.37906, Actual := fbAi.rValue_eu, Delta := 1.0E-3, Message := 'held during glitch');
AssertTrue(Condition := (fbAi.stSts.stCommon.wStatus AND GVL_Const.AI_STS_FAIL_PENDING) <> 0,
           Message := 'fail pending');
fbTime.Advance(tStep := T#100MS);
fbAi(itfTime := fbTime, rIn := 16.0, xChannelFault := FALSE, stCmd := stCmd, stCfg := stCfg);   // после провала
xEverHH := fbAi.xHH;
AssertEquals_REAL(Expected := 52.60415, Actual := fbAi.rValue_eu, Delta := 1.0E-3,
                  Message := 'filter continues from its state (75 if restarted)');
AssertTrue(Condition := fbAi.xValid, Message := 'valid');
FOR iStep := 1 TO 5 DO   // ещё 0,5 с
    fbTime.Advance(tStep := T#100MS);
    fbAi(itfTime := fbTime, rIn := 16.0, stCmd := stCmd, stCfg := stCfg);
    xEverHH := xEverHH OR fbAi.xHH;
END_FOR
AssertFalse(Condition := xEverHH, Message := 'no false HH after a short glitch');
AssertFalse(Condition := fbAi.Fault, Message := 'no failure');

coUnit.TEST_FINISHED();

(* ---- SignalRecoveredClearsFailureAfterDelayAndResetsFilter.method.decl.st ---- *)
// Фильтр 10 с, tFailDelay 2 с: отказ подтверждён; сигнал вернулся (75 %) — отказ держится 1,9 с (значение удерживается
// 50), снимается ровно через 2,0 с, и значение сразу 75: фильтр начался с текущего значения. Без сброса фильтра было бы
// 54,53 (источник: tools/reference/ai_reference.py, сценарий filter «возврат сигнала 50 -> 75 без сброса фильтра»).
METHOD PRIVATE SignalRecoveredClearsFailureAfterDelayAndResetsFilter
VAR
    fbTime : FB_FakeTime;         // подменное время
    fbAi   : FB_AnalogInput;      // ФБ под тестом
    stCmd  : ST_AnalogInputCmd;   // команды
    stCfg  : ST_AnalogInputCfg;   // конфигурация
    iStep  : INT;                 // шаг цикла
END_VAR

(* ---- SignalRecoveredClearsFailureAfterDelayAndResetsFilter.method.impl.st ---- *)
coUnit.TEST('AnalogInput_SignalRecovered_ClearsFailureAfterDelayAndResetsFilter');

stCfg.tFilter := T#10S;
fbAi(itfTime := fbTime, rIn := 12.0, stCmd := stCmd, stCfg := stCfg);   // t0: фильтр начат с 50 %
FOR iStep := 1 TO 30 DO   // обрыв 3 с: отказ подтверждён
    fbTime.Advance(tStep := T#100MS);
    fbAi(itfTime := fbTime, rIn := 0.0, stCmd := stCmd, stCfg := stCfg);
END_FOR
AssertTrue(Condition := fbAi.Fault, Message := 'failure confirmed');
fbTime.Advance(tStep := T#100MS);
fbAi(itfTime := fbTime, rIn := 16.0, stCmd := stCmd, stCfg := stCfg);   // tr: сигнал вернулся, 75 %
FOR iStep := 1 TO 19 DO   // tr + 1,9 с
    fbTime.Advance(tStep := T#100MS);
    fbAi(itfTime := fbTime, rIn := 16.0, stCmd := stCmd, stCfg := stCfg);
END_FOR
AssertTrue(Condition := fbAi.Fault, Message := 'failure kept until tFailDelay after recovery');
AssertFalse(Condition := fbAi.xValid, Message := 'still invalid while recovery is confirmed');
AssertEquals_REAL(Expected := 50.0, Actual := fbAi.rValue_eu, Delta := 1.0E-3, Message := 'value held');
fbTime.Advance(tStep := T#100MS);
fbAi(itfTime := fbTime, rIn := 16.0, stCmd := stCmd, stCfg := stCfg);   // tr + 2,0 с
AssertFalse(Condition := fbAi.Fault, Message := 'failure cleared exactly tFailDelay after recovery');
AssertTrue(Condition := fbAi.xValid, Message := 'valid again');
AssertEquals_REAL(Expected := 75.0, Actual := fbAi.rValue_eu, Delta := 1.0E-3,
                  Message := 'filter restarted from current value (54.53 without restart)');

coUnit.TEST_FINISHED();

(* ---- Sqrt25PctDpReturns50PctFlow.method.decl.st ---- *)
// Корень (расход по перепаду): 8 мА = 25 % перепада — 50 % расхода; 4 мА — 0, 20 мА — 100. источник:
// tools/reference/ai_reference.py, сценарий scale «корень: 8 мА (25 % перепада)».
METHOD PRIVATE Sqrt25PctDpReturns50PctFlow
VAR
    fbTime : FB_FakeTime;         // подменное время
    fbAi   : FB_AnalogInput;      // ФБ под тестом
    stCmd  : ST_AnalogInputCmd;   // команды
    stCfg  : ST_AnalogInputCfg;   // конфигурация
END_VAR

(* ---- StartupWireBreakInvalidUntilFirstGoodValue.method.decl.st ---- *)
// Обрыв уже в первом вызове: удерживать нечего — значение 0.0 и xValid = FALSE сразу (не «годный ноль»), ложного LL
// нет, NE 107 Good до подтверждения; бита AI_STS_FAIL_PENDING нет — значение не удерживается как годное; через 2 с —
// Failure; после возврата и подтверждения — измеренное значение.
METHOD PRIVATE StartupWireBreakInvalidUntilFirstGoodValue
VAR
    fbTime : FB_FakeTime;         // подменное время
    fbAi   : FB_AnalogInput;      // ФБ под тестом
    stCmd  : ST_AnalogInputCmd;   // команды
    stCfg  : ST_AnalogInputCfg;   // конфигурация
    iStep  : INT;                 // шаг цикла
END_VAR

(* ---- StartupWireBreakInvalidUntilFirstGoodValue.method.impl.st ---- *)
coUnit.TEST('AnalogInput_StartupWireBreak_InvalidUntilFirstGoodValue');

stCfg.rRangeHi_eu := 5.0;
SetLimit(stCfgAi := stCfg, uiIdx := E_AiAlarm.LL, xEnable := TRUE, rSp_eu := 0.5, rHyst_eu := 0.1, tOnDly := T#0S,
         tOffDly := T#0S);
fbAi(itfTime := fbTime, rIn := 0.0, stCmd := stCmd, stCfg := stCfg);   // t0: обрыв с первого вызова
AssertFalse(Condition := fbAi.xValid, Message := 'nothing to hold: invalid at once');
AssertEquals_REAL(Expected := 0.0, Actual := fbAi.rValue_eu, Delta := 0.0, Message := 'no good value yet');
AssertFalse(Condition := fbAi.xLL, Message := 'no false LL at startup');
AssertTrue(Condition := fbAi.Status = E_Ne107Status.Good, Message := 'failure not yet confirmed');
AssertTrue(Condition := (fbAi.stSts.stCommon.wStatus AND GVL_Const.AI_STS_FAIL_PENDING) = 0,
           Message := 'no pending bit: nothing is held');
FOR iStep := 1 TO 20 DO   // t0 + 2,0 с
    fbTime.Advance(tStep := T#100MS);
    fbAi(itfTime := fbTime, rIn := 0.0, stCmd := stCmd, stCfg := stCfg);
END_FOR
AssertTrue(Condition := fbAi.Fault, Message := 'failure confirmed');
FOR iStep := 1 TO 1 DO   // tr: сигнал вернулся
    fbTime.Advance(tStep := T#100MS);
    fbAi(itfTime := fbTime, rIn := 16.0, stCmd := stCmd, stCfg := stCfg);
END_FOR
FOR iStep := 1 TO 20 DO   // tr + 2,0 с
    fbTime.Advance(tStep := T#100MS);
    fbAi(itfTime := fbTime, rIn := 16.0, stCmd := stCmd, stCfg := stCfg);
END_FOR
AssertFalse(Condition := fbAi.Fault, Message := 'failure cleared');
AssertTrue(Condition := fbAi.xValid, Message := 'valid');
AssertEquals_REAL(Expected := 3.75, Actual := fbAi.rValue_eu, Delta := 1.0E-5, Message := 'measured value');

coUnit.TEST_FINISHED();

(* ---- SubstitutionDuringFailureLimitsOnSubstValue.method.decl.st ---- *)
// Подмена при подтверждённом отказе датчика (наладка блокировок при оборванной линии): в Manual уставки считаются по
// подменённому значению (11.3, п. 7: принудительный сброс — только в Auto), тревоги уставок подавлены отказом
// (xLimitsOnFail = FALSE), значение годно, NE 107 — Failure. Возврат в Auto при оборванной линии — уставки сняты сразу,
// значение — удерживаемое до отказа, xValid = FALSE.
METHOD PRIVATE SubstitutionDuringFailureLimitsOnSubstValue
VAR
    fbTime : FB_FakeTime;         // подменное время
    fbAi   : FB_AnalogInput;      // ФБ под тестом
    stCmd  : ST_AnalogInputCmd;   // команды
    stCfg  : ST_AnalogInputCfg;   // конфигурация
    iStep  : INT;                 // шаг цикла
    itfAlm : I_Alarm;             // слот тревоги через интерфейс
END_VAR

(* ---- SubstitutionDuringFailureLimitsOnSubstValue.method.impl.st ---- *)
coUnit.TEST('AnalogInput_SubstitutionDuringFailure_LimitsOnSubstValue');

stCfg.tFailDelay := T#1S;
SetLimit(stCfgAi := stCfg, uiIdx := E_AiAlarm.LL, xEnable := TRUE, rSp_eu := 10.0, rHyst_eu := 1.0, tOnDly := T#0S,
         tOffDly := T#0S);
fbAi(itfTime := fbTime, rIn := 12.0, stCmd := stCmd, stCfg := stCfg);   // Auto: 50
FOR iStep := 1 TO 11 DO   // обрыв t0 + 0,1 … t0 + 1,1 с: отказ подтверждён
    fbTime.Advance(tStep := T#100MS);
    fbAi(itfTime := fbTime, rIn := 0.0, stCmd := stCmd, stCfg := stCfg);
END_FOR
AssertTrue(Condition := fbAi.Fault, Message := 'failure confirmed');
AssertFalse(Condition := fbAi.xLL, Message := 'LL forced off in Auto');
stCmd.stCommon.xSetManual := TRUE;
fbTime.Advance(tStep := T#100MS);
fbAi(itfTime := fbTime, rIn := 0.0, stCmd := stCmd, stCfg := stCfg);
AssertTrue(Condition := fbAi.Mode = E_DeviceMode.Manual, Message := 'substitution');
stCmd.rSubstValue_eu := 5.0;   // наладчик проверяет блокировку «сухой ход»
fbTime.Advance(tStep := T#100MS);
fbAi(itfTime := fbTime, rIn := 0.0, stCmd := stCmd, stCfg := stCfg);
AssertEquals_REAL(Expected := 5.0, Actual := fbAi.rValue_eu, Delta := 0.0, Message := 'substituted value');
AssertTrue(Condition := fbAi.xValid, Message := 'substituted value is valid');
AssertTrue(Condition := fbAi.xLL, Message := 'LL on substituted value despite the failure');
AssertTrue(Condition := fbAi.Status = E_Ne107Status.Failure, Message := 'sensor failure still shown');
itfAlm := fbAi.GetAlarm(uiIndex := E_AiAlarm.LL);
AssertTrue(Condition := itfAlm.State = E_AlarmState.SuppressedByDesign, Message := 'LL alarm suppressed by failure');
stCmd.stCommon.xSetAuto := TRUE;
fbTime.Advance(tStep := T#100MS);
fbAi(itfTime := fbTime, rIn := 0.0, stCmd := stCmd, stCfg := stCfg);
AssertFalse(Condition := fbAi.xLL, Message := 'LL forced off again in Auto');
AssertFalse(Condition := fbAi.xValid, Message := 'invalid in Auto with failed sensor');
AssertEquals_REAL(Expected := 50.0, Actual := fbAi.rValue_eu, Delta := 1.0E-4, Message := 'last good value');

coUnit.TEST_FINISHED();

(* ---- SubstitutionNonFiniteValueHeld.method.decl.st ---- *)
// Неконечное значение подмены (NaN с HMI) не принимается: значение остаётся прежним (42), а не NaN.
METHOD PRIVATE SubstitutionNonFiniteValueHeld
VAR
    fbTime : FB_FakeTime;         // подменное время
    fbAi   : FB_AnalogInput;      // ФБ под тестом
    stCmd  : ST_AnalogInputCmd;   // команды
    stCfg  : ST_AnalogInputCfg;   // конфигурация
    uBits  : U_RealBits;          // NaN по битам
END_VAR

(* ---- SubstitutionRenewedAfterTimeoutCountsFullPeriod.method.decl.st ---- *)
// Подмена, снятая по tSubstMax, и новый запрос подмены в следующем же вызове: срок отсчитывается заново,
// подмена не снимается сразу же. Остаток uiSubstRemain_s — целые секунды с округлением вверх
// (59,4 с -> 60, 1,3 с -> 2, 0,1 с -> 1): пока подмена идёт, остаток не 0.
METHOD PRIVATE SubstitutionRenewedAfterTimeoutCountsFullPeriod
VAR
    fbTime : FB_FakeTime;         // подменное время
    fbAi   : FB_AnalogInput;      // ФБ под тестом
    stCmd  : ST_AnalogInputCmd;   // команды
    stCfg  : ST_AnalogInputCfg;   // конфигурация
END_VAR

(* ---- SubstitutionStartsFromCurrentValue.method.decl.st ---- *)
// Слежение: в Auto ФБ пишет rValue_eu в stCmd.rSubstValue_eu, поэтому подмена начинается с текущего значения 7,0 — даже
// если в том же вызове вход изменился (20 мА).
METHOD PRIVATE SubstitutionStartsFromCurrentValue
VAR
    fbTime : FB_FakeTime;         // подменное время
    fbAi   : FB_AnalogInput;      // ФБ под тестом
    stCmd  : ST_AnalogInputCmd;   // команды
    stCfg  : ST_AnalogInputCfg;   // конфигурация
END_VAR

(* ---- SubstitutionTimeoutReturnsToAuto.method.decl.st ---- *)
// tSubstMax 1 мин: подмена 42; остаток uiSubstRemain_s 60 при входе, 1 в 59 с; ровно через 60 с ФБ сам возвращается в
// Auto: результат SubstExpired (+1 к uiCmdSeq), значение измеренное, остаток 0.
METHOD PRIVATE SubstitutionTimeoutReturnsToAuto
VAR
    fbTime : FB_FakeTime;         // подменное время
    fbAi   : FB_AnalogInput;      // ФБ под тестом
    stCmd  : ST_AnalogInputCmd;   // команды
    stCfg  : ST_AnalogInputCfg;   // конфигурация
    iStep  : INT;                 // шаг цикла
    uiSeq  : UINT;                // номер команды до снятия подмены
END_VAR

(* ---- SubstitutionTimeoutReturnsToAuto.method.impl.st ---- *)
coUnit.TEST('AnalogInput_SubstitutionTimeout_ReturnsToAuto');

stCfg.tSubstMax := T#1M;
fbAi(itfTime := fbTime, rIn := 12.0, stCmd := stCmd, stCfg := stCfg);   // Auto: 50
stCmd.stCommon.xSetManual := TRUE;
stCmd.rSubstValue_eu := 42.0;
fbTime.Advance(tStep := T#100MS);
fbAi(itfTime := fbTime, rIn := 12.0, stCmd := stCmd, stCfg := stCfg);   // t0: подмена
AssertEquals_UINT(Expected := 60, Actual := fbAi.stSts.uiSubstRemain_s, Message := '60 s remain at start');
FOR iStep := 1 TO 59 DO   // t0 + 59 с
    fbTime.Advance(tStep := T#1000MS);
    fbAi(itfTime := fbTime, rIn := 12.0, stCmd := stCmd, stCfg := stCfg);
END_FOR
AssertTrue(Condition := fbAi.Mode = E_DeviceMode.Manual, Message := 'still substituted at 59 s');
AssertEquals_REAL(Expected := 42.0, Actual := fbAi.rValue_eu, Delta := 0.0, Message := 'substituted value');
AssertEquals_UINT(Expected := 1, Actual := fbAi.stSts.uiSubstRemain_s, Message := '1 s remains');
uiSeq := fbAi.stSts.stCommon.uiCmdSeq;
fbTime.Advance(tStep := T#1000MS);
fbAi(itfTime := fbTime, rIn := 12.0, stCmd := stCmd, stCfg := stCfg);   // t0 + 60 с
AssertTrue(Condition := fbAi.Mode = E_DeviceMode.Auto, Message := 'back to measurement');
AssertTrue(Condition := fbAi.stSts.stCommon.eCmdResult = E_CmdResult.SubstExpired, Message := 'SubstExpired');
AssertEquals_UINT(Expected := uiSeq + 1, Actual := fbAi.stSts.stCommon.uiCmdSeq, Message := 'counted as one result');
AssertEquals_REAL(Expected := 50.0, Actual := fbAi.rValue_eu, Delta := 1.0E-4, Message := 'measured in the same call');
AssertEquals_UINT(Expected := 0, Actual := fbAi.stSts.uiSubstRemain_s, Message := 'no remaining time');

coUnit.TEST_FINISHED();

(* ---- SubstitutionUnlimitedNoTimeout.method.decl.st ---- *)
// tSubstMax = T#0S — подмена без ограничения срока (Cfg, контракт 11.1): 24 ч в Manual крупными шагами — режим
// остаётся Manual, результата SubstExpired нет, значение подмены, остаток uiSubstRemain_s = 0.
METHOD PRIVATE SubstitutionUnlimitedNoTimeout
VAR
    fbTime : FB_FakeTime;         // подменное время
    fbAi   : FB_AnalogInput;      // ФБ под тестом
    stCmd  : ST_AnalogInputCmd;   // команды
    stCfg  : ST_AnalogInputCfg;   // конфигурация
    iStep  : INT;                 // шаг цикла

    xEverAuto : BOOL;             // режим хоть раз вернулся в Auto
END_VAR

(* ---- SubstitutionUnlimitedNoTimeout.method.impl.st ---- *)
coUnit.TEST('AnalogInput_SubstitutionUnlimited_NoTimeout');

stCfg.tSubstMax := T#0S;
fbAi(itfTime := fbTime, rIn := 12.0, stCmd := stCmd, stCfg := stCfg);
stCmd.stCommon.xSetManual := TRUE;
stCmd.rSubstValue_eu := 42.0;
fbTime.Advance(tStep := T#100MS);
fbAi(itfTime := fbTime, rIn := 12.0, stCmd := stCmd, stCfg := stCfg);                  // подмена
AssertTrue(Condition := fbAi.Mode = E_DeviceMode.Manual, Message := 'substituted');
FOR iStep := 1 TO 24 DO
    fbTime.Advance(tStep := T#1H);
    fbAi(itfTime := fbTime, rIn := 12.0, stCmd := stCmd, stCfg := stCfg);
    xEverAuto := xEverAuto OR fbAi.Mode = E_DeviceMode.Auto;
END_FOR
AssertFalse(Condition := xEverAuto, Message := 'never returned to Auto in 24 h');
AssertTrue(Condition := fbAi.stSts.stCommon.eCmdResult = E_CmdResult.Accepted, Message := 'no SubstExpired');
AssertEquals_REAL(Expected := 42.0, Actual := fbAi.rValue_eu, Delta := 0.0, Message := 'substituted value');
AssertEquals_UINT(Expected := 0, Actual := fbAi.stSts.uiSubstRemain_s, Message := 'no remaining time without a limit');

coUnit.TEST_FINISHED();

(* ---- SubstitutionValueAndCheckFunction.method.decl.st ---- *)
// Подмена (Manual): значение — stCmd.rSubstValue_eu без фильтра, пригодно, NE 107 CheckFunction, бит
// DEV_STS_MODE_MANUAL; уставки считаются по подменённому значению (H 80 при 85). «Измерение» — снова 50.
METHOD PRIVATE SubstitutionValueAndCheckFunction
VAR
    fbTime : FB_FakeTime;         // подменное время
    fbAi   : FB_AnalogInput;      // ФБ под тестом
    stCmd  : ST_AnalogInputCmd;   // команды
    stCfg  : ST_AnalogInputCfg;   // конфигурация
END_VAR

(* ---- SuppressLimitAlarmsInputFlagsStillSet.method.decl.st ---- *)
// xSuppressLimitAlarms: флаг H считается (логика станции его видит), а тревога H — SuppressedByDesign, не
// неквитирована; вход снят — тревога ActiveUnack.
METHOD PRIVATE SuppressLimitAlarmsInputFlagsStillSet
VAR
    fbTime : FB_FakeTime;         // подменное время
    fbAi   : FB_AnalogInput;      // ФБ под тестом
    stCmd  : ST_AnalogInputCmd;   // команды
    stCfg  : ST_AnalogInputCfg;   // конфигурация
    itfAlm : I_Alarm;             // слот тревоги через интерфейс
END_VAR

(* ---- TimeBackwardsFilterHoldsWithoutJump.method.decl.st ---- *)
// «Время назад» (SetNow на 1 с раньше): шаг времени 0 — фильтр стоит, значение не прыгает и конечно; следующий шаг
// вперёд продолжает фильтр от того же значения.
METHOD PRIVATE TimeBackwardsFilterHoldsWithoutJump
VAR
    fbTime  : FB_FakeTime;         // подменное время
    fbAi    : FB_AnalogInput;      // ФБ под тестом
    stCmd   : ST_AnalogInputCmd;   // команды
    stCfg   : ST_AnalogInputCfg;   // конфигурация
    iStep   : INT;                 // шаг цикла
    rBefore : REAL;                // значение до скачка времени
END_VAR

(* ---- TimeBackwardsFilterHoldsWithoutJump.method.impl.st ---- *)
coUnit.TEST('AnalogInput_TimeBackwards_FilterHoldsWithoutJump');

stCfg.tFilter := T#10S;
fbAi(itfTime := fbTime, rIn := 4.0, stCmd := stCmd, stCfg := stCfg);
FOR iStep := 1 TO 50 DO   // 5 с ступени
    fbTime.Advance(tStep := T#100MS);
    fbAi(itfTime := fbTime, rIn := 20.0, stCmd := stCmd, stCfg := stCfg);
END_FOR
rBefore := fbAi.rValue_eu;
fbTime.SetNow(ltValue := fbTime.Now() - LTIME#1S);
fbAi(itfTime := fbTime, rIn := 20.0, stCmd := stCmd, stCfg := stCfg);
AssertEquals_REAL(Expected := rBefore, Actual := fbAi.rValue_eu, Delta := 0.0, Message := 'no jump on time backwards');
AssertTrue(Condition := F_IsFinite(rIn := fbAi.rValue_eu), Message := 'finite');
fbTime.Advance(tStep := T#100MS);
fbAi(itfTime := fbTime, rIn := 20.0, stCmd := stCmd, stCfg := stCfg);
AssertTrue(Condition := fbAi.rValue_eu > rBefore, Message := 'filter continues forward');
AssertTrue(Condition := fbAi.rValue_eu < rBefore + 1.0, Message := 'by one 100 ms step only');

coUnit.TEST_FINISHED();

(* ---- WireBreakHoldsLastGoodValue.method.decl.st ---- *)
// HoldLast (по умолчанию): при обрыве значение 3,75 (16 мА на шкале 0..5) держится и до подтверждения, и после него
// (xValid = FALSE); проценты и слежение в stCmd — то же значение.
METHOD PRIVATE WireBreakHoldsLastGoodValue
VAR
    fbTime : FB_FakeTime;         // подменное время
    fbAi   : FB_AnalogInput;      // ФБ под тестом
    stCmd  : ST_AnalogInputCmd;   // команды
    stCfg  : ST_AnalogInputCfg;   // конфигурация
    iStep  : INT;                 // шаг цикла
END_VAR

(* ---- WireBreakHoldsLastGoodValue.method.impl.st ---- *)
coUnit.TEST('AnalogInput_WireBreak_HoldsLastGoodValue');

stCfg.rRangeHi_eu := 5.0;
fbAi(itfTime := fbTime, rIn := 16.0, stCmd := stCmd, stCfg := stCfg);   // t0: 75 % = 3,75
FOR iStep := 1 TO 10 DO   // обрыв, t0 + 1,0 с
    fbTime.Advance(tStep := T#100MS);
    fbAi(itfTime := fbTime, rIn := 0.0, stCmd := stCmd, stCfg := stCfg);
END_FOR
AssertEquals_REAL(Expected := 3.75, Actual := fbAi.rValue_eu, Delta := 1.0E-5, Message := 'held while pending');
FOR iStep := 1 TO 20 DO   // t0 + 3,0 с: отказ подтверждён
    fbTime.Advance(tStep := T#100MS);
    fbAi(itfTime := fbTime, rIn := 0.0, stCmd := stCmd, stCfg := stCfg);
END_FOR
AssertTrue(Condition := fbAi.Fault, Message := 'failure confirmed');
AssertEquals_REAL(Expected := 3.75, Actual := fbAi.rValue_eu, Delta := 1.0E-5, Message := 'held after confirmation');
AssertEquals_REAL(Expected := 75.0, Actual := fbAi.rValue_pct, Delta := 1.0E-4, Message := 'percent of held value');
AssertEquals_REAL(Expected := 3.75, Actual := stCmd.rSubstValue_eu, Delta := 0.0, Message := 'tracking of held value');
AssertFalse(Condition := fbAi.xValid, Message := 'held value is not valid');

coUnit.TEST_FINISHED();

(* ---- WireBreakSetsFailureAfterDelay.method.decl.st ---- *)
// Обрыв (0 мА) при tFailDelay = 2 с: до 1,9 с отказа нет, значение удерживается (2,5 м), ложного LL нет, бит
// AI_STS_FAIL_PENDING; ровно через 2,0 с — Failure, xValid = FALSE, бит AI_FLT_FAIL_LOW (AI_STS_FAIL_PENDING снят),
// тревога Failure, LL снят принудительно. Образец — раздел 23.3 контракта.
METHOD PRIVATE WireBreakSetsFailureAfterDelay
VAR
    fbTime : FB_FakeTime;         // подменное время
    fbAi   : FB_AnalogInput;      // ФБ под тестом
    stCmd  : ST_AnalogInputCmd;   // команды
    stCfg  : ST_AnalogInputCfg;   // конфигурация
    itfAlm : I_Alarm;             // слот тревоги через интерфейс
    iStep  : INT;                 // шаг цикла
END_VAR

(* ---- WireBreakSetsFailureAfterDelay.method.impl.st ---- *)
coUnit.TEST('AnalogInput_WireBreak_SetsFailureAfterDelay');

stCfg.rRangeHi_eu := 5.0;
SetLimit(stCfgAi := stCfg, uiIdx := E_AiAlarm.LL, xEnable := TRUE, rSp_eu := 0.5, rHyst_eu := 0.0, tOnDly := T#0S,
         tOffDly := T#0S);
fbAi(itfTime := fbTime, rIn := 12.0, stCmd := stCmd, stCfg := stCfg);   // t0: 50 % = 2,5 м
fbTime.Advance(tStep := T#100MS);
fbAi(itfTime := fbTime, rIn := 0.0, stCmd := stCmd, stCfg := stCfg);   // t1 = t0 + 0,1 с: обрыв
FOR iStep := 1 TO 19 DO   // t1 + 1,9 с
    fbTime.Advance(tStep := T#100MS);
    fbAi(itfTime := fbTime, rIn := 0.0, stCmd := stCmd, stCfg := stCfg);
END_FOR
AssertFalse(Condition := fbAi.Fault, Message := 'no failure before tFailDelay');
AssertEquals_REAL(Expected := 2.5, Actual := fbAi.rValue_eu, Delta := 1.0E-4, Message := 'last good value held');
AssertFalse(Condition := fbAi.xLL, Message := 'no false LL on wire break');
AssertTrue(Condition := fbAi.xValid, Message := 'value still valid while failure is pending');
AssertTrue(Condition := (fbAi.stSts.stCommon.wStatus AND GVL_Const.AI_STS_FAIL_PENDING) <> 0,
           Message := 'fail pending bit');
AssertTrue(Condition := fbAi.stSts.eSignal = E_AiSignalState.FailLow, Message := 'instant classification FailLow');
fbTime.Advance(tStep := T#100MS);
fbAi(itfTime := fbTime, rIn := 0.0, stCmd := stCmd, stCfg := stCfg);   // t1 + 2,0 с
AssertTrue(Condition := fbAi.Status = E_Ne107Status.Failure, Message := 'failure after 2 s');
AssertFalse(Condition := fbAi.xValid, Message := 'value invalid after confirmed failure');
AssertEquals_WORD(Expected := GVL_Const.AI_FLT_FAIL_LOW, Actual := fbAi.stSts.stCommon.wFault,
                  Message := 'fault bit FAIL_LOW');
AssertTrue(Condition := (fbAi.stSts.stCommon.wStatus AND GVL_Const.AI_STS_SIGNAL_FAIL) <> 0, Message := 'fail bit');
AssertTrue(Condition := (fbAi.stSts.stCommon.wStatus AND GVL_Const.AI_STS_FAIL_PENDING) = 0,
           Message := 'pending bit cleared after confirmation');
AssertFalse(Condition := fbAi.xLL, Message := 'LL forced off on failure');
itfAlm := fbAi.GetAlarm(uiIndex := E_AiAlarm.Failure);
AssertTrue(Condition := itfAlm.State = E_AlarmState.ActiveUnack, Message := 'failure alarm annunciated');

coUnit.TEST_FINISHED();

(* ---- WireBreakShorterThanDelayNoFailure.method.decl.st ---- *)
// Обрыв на 1,5 с при tFailDelay = 2 с: отказа и тревоги нет ни в одном вызове, значение держится, после возврата
// сигнала — сразу новое измеренное значение; ещё 3 с — без отказа.
METHOD PRIVATE WireBreakShorterThanDelayNoFailure
VAR
    fbTime     : FB_FakeTime;         // подменное время
    fbAi       : FB_AnalogInput;      // ФБ под тестом
    stCmd      : ST_AnalogInputCmd;   // команды
    stCfg      : ST_AnalogInputCfg;   // конфигурация
    itfAlm     : I_Alarm;             // слот тревоги через интерфейс
    iStep      : INT;                 // шаг цикла
    xEverFault : BOOL;                // отказ был хотя бы в одном вызове
END_VAR

(* ---- WireBreakShorterThanDelayNoFailure.method.impl.st ---- *)
coUnit.TEST('AnalogInput_WireBreakShorterThanDelay_NoFailure');

stCfg.rRangeHi_eu := 5.0;
fbAi(itfTime := fbTime, rIn := 12.0, stCmd := stCmd, stCfg := stCfg);   // t0: 2,5
FOR iStep := 1 TO 15 DO                                           // обрыв t0 + 0,1 … t0 + 1,5 с
    fbTime.Advance(tStep := T#100MS);
    fbAi(itfTime := fbTime, rIn := 0.0, stCmd := stCmd, stCfg := stCfg);
    xEverFault := xEverFault OR fbAi.Fault OR NOT fbAi.xValid;
END_FOR
AssertEquals_REAL(Expected := 2.5, Actual := fbAi.rValue_eu, Delta := 1.0E-4, Message := 'held during short break');
FOR iStep := 1 TO 30 DO                                           // сигнал вернулся: 16 мА, 3 с
    fbTime.Advance(tStep := T#100MS);
    fbAi(itfTime := fbTime, rIn := 16.0, stCmd := stCmd, stCfg := stCfg);
    xEverFault := xEverFault OR fbAi.Fault OR NOT fbAi.xValid;
END_FOR
AssertFalse(Condition := xEverFault, Message := 'break shorter than tFailDelay gives no failure');
AssertEquals_REAL(Expected := 3.75, Actual := fbAi.rValue_eu, Delta := 1.0E-5, Message := 'measured after return');
itfAlm := fbAi.GetAlarm(uiIndex := E_AiAlarm.Failure);
AssertTrue(Condition := itfAlm.State = E_AlarmState.Normal, Message := 'no failure alarm');

coUnit.TEST_FINISHED();
